TYPE "DT_DIGITAL_INPUT_MIV_AND_BYPASS"
VERSION : 0.1
   STRUCT
      MIV_CLOSED { S7_SetPoint := 'False'} : "DT_STATUS_SOLO" := ((FALSE, 1, 192), (32000, 32000, 32000), (0, 1, 4), (FALSE, FALSE, 0));
      MIV_INTERMEDIATE { S7_SetPoint := 'False'} : "DT_STATUS_SOLO" := ((FALSE, 1, 193), (32000, 32000, 32000), (0, 0, 0), (FALSE, FALSE, 0));
      MIV_OPEN { S7_SetPoint := 'False'} : "DT_STATUS_SOLO" := ((FALSE, 1, 194), (32000, 32000, 32000), (0, 1, 4), (FALSE, FALSE, 0));
      MIV_SAFETY_PIN { S7_SetPoint := 'False'} : "DT_STATUS_SOLO" := ((FALSE, 1, 195), (32000, 32000, 32000), (0, 0, 0), (FALSE, FALSE, 0));
      MIV_FILLING_POSITION { S7_SetPoint := 'False'} : "DT_STATUS_SOLO" := ((FALSE, 1, 196), (32000, 32000, 32000), (0, 0, 0), (FALSE, FALSE, 0));
      MIV_MCB_ON { S7_SetPoint := 'False'} : "DT_STATUS_SOLO" := ((FALSE, 1, 197), (32000, 32000, 32000), (0, 3, 4), (FALSE, FALSE, 0));
      MIV_CONT_ON { S7_SetPoint := 'False'} : "DT_STATUS_SOLO" := ((FALSE, 1, 198), (32000, 32000, 32000), (0, 1, 4), (FALSE, FALSE, 0));
      MIV_HEATER_MCB_OK { S7_SetPoint := 'False'} : "DT_STATUS_SOLO" := ((FALSE, 1, 199), (32000, 32000, 32000), (0, 3, 4), (FALSE, FALSE, 0));
      SPARE_200 { S7_SetPoint := 'False'} : "DT_STATUS_SOLO" := ((FALSE, 1, 200), (32000, 32000, 32000), (0, 0, 0), (FALSE, FALSE, 0));
      BYPASS_OPEN { S7_SetPoint := 'False'} : "DT_STATUS_SOLO" := ((FALSE, 1, 201), (32000, 32000, 32000), (0, 1, 4), (FALSE, FALSE, 0));
      BYPASS_CLOSED { S7_SetPoint := 'False'} : "DT_STATUS_SOLO" := ((FALSE, 1, 202), (32000, 32000, 32000), (0, 1, 4), (FALSE, FALSE, 0));
      BYPASS_MCB_ON { S7_SetPoint := 'False'} : "DT_STATUS_SOLO" := ((FALSE, 1, 203), (32000, 32000, 32000), (0, 3, 4), (FALSE, FALSE, 0));
      BYPASS_MCB_TRIP { S7_SetPoint := 'False'} : "DT_STATUS_SOLO" := ((FALSE, 1, 204), (32000, 32000, 32000), (0, 0, 0), (FALSE, FALSE, 0));
      BYPASS_CONT_ON { S7_SetPoint := 'False'} : "DT_STATUS_SOLO" := ((FALSE, 1, 205), (32000, 32000, 32000), (0, 0, 0), (FALSE, FALSE, 0));
      BYPASS_CONT_OPEN_ON { S7_SetPoint := 'False'} : "DT_STATUS_SOLO" := ((FALSE, 1, 206), (32000, 32000, 32000), (0, 1, 4), (FALSE, FALSE, 0));
      BYPASS_CONT_CLOSE_ON { S7_SetPoint := 'False'} : "DT_STATUS_SOLO" := ((FALSE, 1, 207), (32000, 32000, 32000), (0, 1, 4), (FALSE, FALSE, 0));
      BYPASS_TORQUE_OPEN_OK { S7_SetPoint := 'False'} : "DT_STATUS_SOLO" := ((FALSE, 1, 208), (32000, 32000, 32000), (0, 1, 3), (FALSE, FALSE, 0));
      BYPASS_TORQUE_CLOSE_OK { S7_SetPoint := 'False'} : "DT_STATUS_SOLO" := ((FALSE, 1, 209), (32000, 32000, 32000), (0, 0, 0), (FALSE, FALSE, 0));
      BYPASS_THERMAL_OVERLOAD { S7_SetPoint := 'False'} : "DT_STATUS_SOLO" := ((FALSE, 1, 210), (32000, 32000, 32000), (0, 0, 0), (FALSE, FALSE, 0));
      BYPASS_HEATER_MCB_OK { S7_SetPoint := 'False'} : "DT_STATUS_SOLO" := ((FALSE, 1, 211), (32000, 32000, 32000), (0, 0, 0), (FALSE, FALSE, 0));
      BYPASS_FAULT { S7_SetPoint := 'False'} : "DT_STATUS_SOLO" := ((FALSE, 1, 212), (32000, 32000, 32000), (0, 0, 0), (FALSE, FALSE, 0));
      MCB_Trip { S7_SetPoint := 'False'} : "DT_STATUS_SOLO" := ((FALSE, 1, 213), (32000, 32000, 32000), (0, 0, 0), (FALSE, FALSE, 0));
      MIV_TORQUE_CLOSED { S7_SetPoint := 'False'} : "DT_STATUS_SOLO" := ((FALSE, 1, 214), (32000, 32000, 32000), (0, 1, 4), (FALSE, FALSE, 0));
      MIV_TORQUE_OPEN { S7_SetPoint := 'False'} : "DT_STATUS_SOLO" := ((FALSE, 1, 215), (32000, 32000, 32000), (0, 1, 4), (FALSE, FALSE, 0));
      MIV_THERMOSWITCH { S7_SetPoint := 'False'} : "DT_STATUS_SOLO" := ((FALSE, 1, 216), (32000, 32000, 32000), (0, 4, 3), (FALSE, FALSE, 0));
      SPARE_217 { S7_SetPoint := 'False'} : "DT_STATUS_SOLO" := ((FALSE, 1, 217), (32000, 32000, 32000), (0, 0, 0), (FALSE, FALSE, 0));
      SPARE_218 { S7_SetPoint := 'False'} : "DT_STATUS_SOLO" := ((FALSE, 1, 218), (32000, 32000, 32000), (0, 0, 0), (FALSE, FALSE, 0));
      SPARE_219 { S7_SetPoint := 'False'} : "DT_STATUS_SOLO" := ((FALSE, 1, 219), (32000, 32000, 32000), (0, 0, 0), (FALSE, FALSE, 0));
      SPARE_220 { S7_SetPoint := 'False'} : "DT_STATUS_SOLO" := ((FALSE, 1, 220), (32000, 32000, 32000), (0, 0, 0), (FALSE, FALSE, 0));
      SPARE_221 { S7_SetPoint := 'False'} : "DT_STATUS_SOLO" := ((FALSE, 1, 221), (32000, 32000, 32000), (0, 0, 0), (FALSE, FALSE, 0));
      SPARE_222 { S7_SetPoint := 'False'} : "DT_STATUS_SOLO" := ((FALSE, 1, 222), (32000, 32000, 32000), (0, 0, 0), (FALSE, FALSE, 0));
      SPARE_223 { S7_SetPoint := 'False'} : "DT_STATUS_SOLO" := ((FALSE, 1, 223), (32000, 32000, 32000), (0, 0, 0), (FALSE, FALSE, 0));
   END_STRUCT;

END_TYPE

